(* IEC 61131-3 sources: repolevel_ST_code_completion/output/0122完整版本_无planner目前sota/repoeval_Wrappers/readful_result, 1 file *)

(* ---- FB_Wrapper.st ---- *)
FUNCTION_BLOCK FB_Wrapper
VAR_INPUT
	in:BOOL;
END_VAR
VAR_OUTPUT
	out:BOOL;
END_VAR
<UNFIXABLE>
END_FUNCTION_BLOCK
